// // MIGRATION DRAFT: not included in PLC compilation.
// // Reference: Reference_Project/GateAccess_Station_FB.scl, object GateAccess_Station_FB.
// // Types, globals, calls, units and behavior require manual reconciliation.
// // See docs/TIA_Missing_Blocks.md before importing as PLC code.
// // SAFETY REVIEW REQUIRED: not a TwinSAFE implementation.
FUNCTION_BLOCK GateAccess_Station_FB
// 
//    VAR_INPUT
//       Sys_No : UInt;
//       Right_True   : Bool;
//       Switches   : Byte;
//       GateLockedFeedback : Bool;
//       NoEStop : Bool;
//       I_G1_GuardOpen : Bool;
//       I_L1_Unlocked : Bool;
//       FaultResetCmd : Bool;
//       AllDrivesHealthy : Bool;
//       SafetyResetDone : Bool;
//       NoVTDLocalMode : Bool;
//       NoCrossoverPaused : Bool;
//       Safe_Bypassed : Bool;
//       LGX_Secure_Access : Bool;
//       AllDevicesStopped : Bool;
//    END_VAR
// 
//    VAR_OUTPUT
//       Lamps   : Byte;
//       O_S1_SolenoidEnergise : Bool;
//       Lock_Reset   : Bool;
//       CurrentState : UInt;
//       GateFault : Bool;
//    END_VAR
// 
//    VAR_IN_OUT
//       Gate_Station : Gate_Station_UDT;
//    END_VAR
// 
//    VAR
//       RTE_PB : Bool;
//       Reset_PB : Bool;
//       Restart_PB : Bool;
//       GateAccessControl   : GateAccessControl_FB;
//       ModeManager   : ModeManager_FB;
//    END_VAR
// 
//    VAR_TEMP
//       i : UInt;
//    END_VAR
// 
//    VAR CONSTANT
//       AUTO_RUNNING : UInt := 0;
//       RTE_REQUESTED : UInt := 1;
//       SAFE_TO_UNLOCK : UInt := 3;
//       ACCESS_MANUAL_MODE : UInt := 4;
//       RESETTING : UInt := 6;
//    END_VAR

// // MIGRATION DRAFT: not included in PLC compilation.
// // Reference: Reference_Project/GateAccess_Station_FB.scl, object GateAccess_Station_FB.
// // Types, globals, calls, units and behavior require manual reconciliation.
// // See docs/TIA_Missing_Blocks.md before importing as PLC code.
// // SAFETY REVIEW REQUIRED: not a TwinSAFE implementation.
// IF Right_True THEN
// 
// 	    Reset_PB := Switches.%X1;
// 	    Restart_PB := Switches.%X3;
// 	    RTE_PB := Switches.%X2;
// 	ELSE
// 
// 	    Restart_PB := Switches.%X3;
// 	    Reset_PB := Switches.%X2;
// 	    RTE_PB := Switches.%X1;
// 	END_IF;
// 
// 	GateAccessControl(
// 	                   UnlockPermissive := ModeManager.GateUnlockPermissive,
// 	                   FaultResetCmd := FaultResetCmd,
// 	                   I_G1_GuardOpen := I_G1_GuardOpen,
// 	                   I_L1_Unlocked := I_L1_Unlocked,
// 	                   GateLockedFeedback := GateLockedFeedback,
// 	                   NoEStop := NoEStop
// 	);
// 
// 	ModeManager(
// 	             RTE_PB := RTE_PB,
// 	             Reset_PB := Reset_PB,
// 	             Restart_PB := Restart_PB,
// 	             GateClosed := GateAccessControl.GateClosed,
// 	             GateLockedFeedback := GateLockedFeedback,
// 	             GateFault := GateAccessControl.GateFault,
// 	             NoEStop := NoEStop,
// 	             AllDrivesHealthy := AllDrivesHealthy,
// 	             SafetyResetDone := SafetyResetDone,
// 	             NoVTDLocalMode := NoVTDLocalMode,
// 	             NoCrossoverPaused := NoCrossoverPaused,
// 	             AllDevicesStopped := Gate_Station.Secure_Access AND AllDevicesStopped AND LGX_Secure_Access,
// 	             Safe_Bypassed := Safe_Bypassed,
// 	             ForceRTE := GateAccessControl.ForceRTE_Request,
// 	             Reset := FaultResetCmd
// 	);
// 
// 	O_S1_SolenoidEnergise := GateAccessControl.O_S1_SolenoidEnergise;
// 	CurrentState := ModeManager.CurrentState;
// 	GateFault := GateAccessControl.GateFault;
// 
// 	IF ModeManager.CurrentState = RESETTING AND Sys_No <> 0 THEN
// 	    FOR i := Settings_DB.VTD[Sys_No].Lowest_Level TO Settings_DB.VTD[Sys_No].Highest_Level DO
// 	        Control.VTD[Sys_No].Instruction.Reset :=
// 	        Control.ECnv_Sys[Sys_No].Instruction.Reset :=
// 	        Control.LCnv_Sys[Sys_No].Cnv_Level[i].Cnv1.Instruction.Reset :=
// 	        Control.LCnv_Sys[Sys_No].Cnv_Level[i].Cnv2.Instruction.Reset := TRUE;
// 	    END_FOR;
// 
// 	    IF AllDrivesHealthy THEN
// 	        FOR i := Settings_DB.VTD[Sys_No].Lowest_Level TO Settings_DB.VTD[Sys_No].Highest_Level DO
// 	            Control.VTD[Sys_No].Instruction.Reset :=
// 	            Control.ECnv_Sys[Sys_No].Instruction.Reset :=
// 	            Control.LCnv_Sys[Sys_No].Cnv_Level[i].Cnv1.Instruction.Reset :=
// 	            Control.LCnv_Sys[Sys_No].Cnv_Level[i].Cnv2.Instruction.Reset := FALSE;
// 	        END_FOR;
// 
// 	        FOR i := Settings_DB.VTD[Sys_No].Lowest_Level TO Settings_DB.VTD[Sys_No].Highest_Level DO
// 	            Control.VTD[Sys_No].Instruction.Mode_Change :=
// 	            Control.ECnv_Sys[Sys_No].Instruction.Mode_Change :=
// 	            Control.LCnv_Sys[Sys_No].Cnv_Level[i].Cnv1.Instruction.Mode_Change :=
// 	            Control.LCnv_Sys[Sys_No].Cnv_Level[i].Cnv2.Instruction.Mode_Change :=
// 	            Control.LCnv_Sys[Sys_No].Cnv_Level[i].Cnv1.Safety_Stop_Cnrl.Mode :=
// 	            Control.LCnv_Sys[Sys_No].Cnv_Level[i].Cnv2.Safety_Stop_Cnrl.Mode := 3;
// 
// 	            Control.VTD[Sys_No].Instruction.Enable :=
// 	            Control.ECnv_Sys[Sys_No].Instruction.Enable :=
// 	            Control.LCnv_Sys[Sys_No].Cnv_Level[i].Cnv1.Instruction.Enable :=
// 	            Control.LCnv_Sys[Sys_No].Cnv_Level[i].Cnv2.Instruction.Enable := TRUE;
// 	        END_FOR;
// 	    END_IF;
// 	END_IF;
// 
// 
// 	IF ModeManager.CurrentState = ACCESS_MANUAL_MODE AND Sys_No <> 0 THEN
// 	    FOR i := Settings_DB.VTD[Sys_No].Lowest_Level TO Settings_DB.VTD[Sys_No].Highest_Level DO
// 	        Control.VTD[Sys_No].Instruction.Mode_Change :=
// 	        Control.ECnv_Sys[Sys_No].Instruction.Mode_Change :=
// 	        Control.LCnv_Sys[Sys_No].Cnv_Level[i].Cnv1.Instruction.Mode_Change :=
// 	        Control.LCnv_Sys[Sys_No].Cnv_Level[i].Cnv2.Instruction.Mode_Change :=
// 	        Control.LCnv_Sys[Sys_No].Cnv_Level[i].Cnv1.Safety_Stop_Cnrl.Mode :=
// 	        Control.LCnv_Sys[Sys_No].Cnv_Level[i].Cnv2.Safety_Stop_Cnrl.Mode := 1;
// 	    END_FOR;
// 	END_IF;
// 
// 	IF Right_True THEN
// 	    Lamps.%X0 := (NOT NoEStop OR GateAccessControl.GateFault) AND Clock_1Hz;
// 	    Lamps.%X3 := (ModeManager.ReqFlash_RestartLamp AND Clock_1Hz) OR ModeManager.RestartLampSteadyOn;
// 	    Lamps.%X1 := ModeManager.ReqFlash_ResetLamp AND Clock_1Hz;
// 	    Lamps.%X2 := ModeManager.ReqFlash_RTE_Lamp OR (ModeManager.CurrentState = SAFE_TO_UNLOCK AND NOT NoEStop) OR ModeManager.CurrentState = SAFE_TO_UNLOCK OR ModeManager.CurrentState = ACCESS_MANUAL_MODE;
// 	ELSE
// 	    Lamps.%X0 := (NOT NoEStop OR GateAccessControl.GateFault) AND Clock_1Hz;
// 	    Lamps.%X2 := ModeManager.ReqFlash_ResetLamp AND Clock_1Hz;
// 	    Lamps.%X3 := (ModeManager.ReqFlash_RestartLamp AND Clock_1Hz) OR ModeManager.RestartLampSteadyOn;
// 	    Lamps.%X1 := ModeManager.ReqFlash_RTE_Lamp OR (ModeManager.CurrentState = SAFE_TO_UNLOCK AND NOT NoEStop) OR ModeManager.CurrentState = SAFE_TO_UNLOCK OR ModeManager.CurrentState = ACCESS_MANUAL_MODE;
// 	END_IF;
// 
// 
// 
// 	Gate_Station.Requested_Access := ModeManager.CurrentState = RTE_REQUESTED;
// 	Gate_Station.Safe_To_Restart := ModeManager.RestartLampSteadyOn;

END_FUNCTION_BLOCK

(* stored: Version 1.1.0.1
   POU GateAccess_Station_FB: Id {3205d1a7-4fed-5a02-a09a-24417c3de077}, SpecialFunc None *)
